// TwinCAT 3 PLC project SendData
// ProgramVersion: 3.1.4023.0
// libraries:
//   Tc2_Standard, * (Beckhoff Automation GmbH)
//   Tc2_System, * (Beckhoff Automation GmbH)
//   Tc3_Module, * (Beckhoff Automation GmbH)
// project tree:
//   / PlcTask.TcTTO
//   POUs/ MAIN.TcPOU
// real-time tasks:
//   TASK PlcTask: cycle T#10ms, priority 20, ADS port 350
// I/O:
//   DEVICE Device 2 (EtherCAT), AmsNetId 192.168.18.191.3.1
//     Box 1 (sample_app) [sample_app]
//     Box 2 (sample_app) [sample_app]
// variable links:
//   SendData/SendData Instance <-> Device 2 (EtherCAT)/Box 1 (sample_app)
//     PlcTask Inputs/MAIN.rawAngleM1 <-> Inputs process data mapping/Counter
//     PlcTask Outputs/MAIN.dummyDataM1 <-> Outputs process data mapping/Trigger
//   SendData/SendData Instance <-> Device 2 (EtherCAT)/Box 2 (sample_app)
//     PlcTask Inputs/MAIN.rawAngleM2 <-> Inputs process data mapping/Counter
//     PlcTask Outputs/MAIN.dummyDataM2 <-> Outputs process data mapping/Trigger

CONFIGURATION SendData
    RESOURCE PLC ON TwinCAT3
        TASK PlcTask(INTERVAL := T#10ms, PRIORITY := 20);
        PROGRAM MAIN WITH PlcTask : MAIN;
    END_RESOURCE
END_CONFIGURATION

// ---- POUs/MAIN.TcPOU
PROGRAM MAIN
VAR
	dirM1 : BYTE := 1;
	speedM1 : WORD := 100;
	dummyDataM1 AT %Q*: DWORD := SHL(dirM1,2*8) OR speedM1 ;
	rawAngleM1 AT %I*: DWORD;
	angleM1: REAL;
	
	dirM2 : BYTE := 1;
	speedM2 : WORD := 100;
	dummyDataM2 AT %Q*: DWORD := SHL(dirM2,2*8) OR speedM2 ;
	rawAngleM2 AT %I*: DWORD;
	angleM2: REAL;
END_VAR

dummyDataM1 := SHL(dirM1,2*8) OR speedM1 ;
angleM1 := (rawAngleM1/100.0) - 180;
dummyDataM2 := SHL(dirM2,2*8) OR speedM2 ;
angleM2 := (rawAngleM2/100.0) - 180;
speedM2 := speedM1/2;

END_PROGRAM
